TYPE tea :
STRUCT

price			: REAL;
name			: STRING;
ingredients		: STRING;	


END_STRUCT
END_TYPE

(* stored: Version 1.1.0.1
   DUT tea: Id {4e6c541a-3b84-4a53-937a-8e596cb94f94} *)
